(* IEC 61131-3 sources: SRCI_CLIENT_PLC/RobotLibrary/Library/Structures/Telegram/RobToPlc/Sequence, 2 files *)

(* ---- TelegramRobToPlcSequence.st ---- *)
{attribute 'pack_mode' := '1'}
// -------------------------------------------------------------------------
//  SRCI Robot Library
// -------------------------------------------------------------------------
//
//  Object:      TelegramPlcToRobSequence
//  Author:      Thorsten Brach
//  Date:        2024-11-02
//
//  Description:
//
//
//  Copyright:
//    (C) 2024 Thorsten Brach. All rights reserved
//             Licensed under the MIT License.
//
//  Disclaimer:
//    This project is provided without any guarantee and can be used for
//    private and commercial purposes. Any use is at the user’s
//    own risk and responsibility.
//
// -------------------------------------------------------------------------
TYPE TelegramRobToPlcSequence :
STRUCT
  /// Header
  Header   : TelegramRobToPlcSequenceHeader;
  /// Fragment
  Fragment : ARRAY[0..RobotLibraryParameter.FRAGMENT_MAX] OF TelegramRobToPlcFragment;
END_STRUCT
END_TYPE

(* ---- TelegramRobToPlcSequenceHeader.st ---- *)
{attribute 'pack_mode' := '1'}
// -------------------------------------------------------------------------
//  SRCI Robot Library
// -------------------------------------------------------------------------
//
//  Object:      TelegramRobToPlcSequenceHeader
//  Author:      Thorsten Brach
//  Date:        2024-11-02
//
//  Description:
//
//
//  Copyright:
//    (C) 2024 Thorsten Brach. All rights reserved
//             Licensed under the MIT License.
//
//  Disclaimer:
//    This project is provided without any guarantee and can be used for
//    private and commercial purposes. Any use is at the user’s
//    own risk and responsibility.
//
// -------------------------------------------------------------------------
TYPE TelegramRobToPlcSequenceHeader :
STRUCT
  /// Telegram Sequence and Acknowledgement number
  SEQ_ACK      : UINT;
  /// Length of the Telegram Sequence excluding this Telegram Sequence Header
  PayloadLength : UINT;
END_STRUCT
END_TYPE
